Fanuc KAREL source: kt00731.KL

-- PROVISIONAL review KL for V770-1; original PC SHA256 601eb702e2eab291c6392ab3cd3199fc0efa8b6afa8decdce22468af8dde6592
-- Incomplete behavior may be omitted. Consult companion uncertainty JSON. Do not deploy.
PROGRAM KT00731
%NOLOCKGROUP
VAR
  OUT : INTEGER
-- UNRESOLVED_DECL ARG type=002010
BEGIN
  -- UNRESOLVED_PC offsets 5-18; opcodes 22,1D,23
  -- UNRESOLVED_PC offsets 23-27; opcodes 7F
END KT00731
